(* IEC 61131-3 sources: llm-plc-st-eval/data/definitivo/gemini-3.1-pro-preview/I8/few_shot, 3 files *)

(* ---- ejec_1.st ---- *)
FUNCTION_BLOCK FB_Compresor
VAR_INPUT
    pOilOk : BOOL;    (* Presion de aceite correcta *)
    tempOk : BOOL;    (* Temperatura correcta *)
    sinAlm : BOOL;    (* Ausencia de alarmas *)
    btnMarcha : BOOL; (* Boton de arranque *)
    btnParo : BOOL;   (* Boton de parada *)
END_VAR
VAR_OUTPUT
    comp : BOOL;      (* Salida del compresor *)
    causaBloqueo : INT; (* Causa de bloqueo: 1=Aceite, 2=Temp, 3=Alarma, 0=Ninguno *)
END_VAR
VAR
    tonOil : TON;     (* Temporizador para presion de aceite *)
    trigMarcha : R_TRIG; (* Detector de flanco para boton de marcha *)
    permisivosOk : BOOL; (* Estado de todos los permisivos *)
END_VAR

(* Temporizador: presion de aceite activa por 3 segundos continuos *)
tonOil(IN := pOilOk, PT := T#3S);

(* Determinacion de la causa de bloqueo con prioridad (menor numero primero) *)
IF NOT tonOil.Q THEN
    causaBloqueo := 1;
ELSIF NOT tempOk THEN
    causaBloqueo := 2;
ELSIF NOT sinAlm THEN
    causaBloqueo := 3;
ELSE
    causaBloqueo := 0;
END_IF;

(* Evaluacion global de permisivos *)
permisivosOk := (causaBloqueo = 0);

(* Deteccion de flanco de subida del boton de marcha *)
trigMarcha(CLK := btnMarcha);

(* Logica de control del compresor (Paro prioritario y perdida de permisivos) *)
IF btnParo OR NOT permisivosOk THEN
    comp := FALSE;
ELSIF trigMarcha.Q AND permisivosOk THEN
    comp := TRUE;
END_IF;
END_FUNCTION_BLOCK

(* ---- ejec_2.st ---- *)
FUNCTION_BLOCK FB_Compresor
VAR_INPUT
    pOilOk : BOOL; (* Presion de aceite *)
    tempOk : BOOL; (* Temperatura correcta *)
    sinAlm : BOOL; (* Ausencia de alarmas *)
    btnMarcha : BOOL; (* Boton de arranque *)
    btnParo : BOOL; (* Boton de parada *)
END_VAR
VAR_OUTPUT
    comp : BOOL; (* Mando del compresor *)
    causaBloqueo : INT; (* Codigo de permisivo faltante *)
END_VAR
VAR
    tOil : TON; (* Temporizador de presion de aceite *)
    trigMarcha : R_TRIG; (* Detector de flanco de marcha *)
    permisivosOk : BOOL; (* Estado de todos los permisivos *)
END_VAR

(* Temporizador para validar la presion de aceite por 3s continuos *)
tOil(IN := pOilOk, PT := T#3S);

(* Deteccion de flanco de subida del boton de marcha *)
trigMarcha(CLK := btnMarcha);

(* Evaluacion general de permisivos *)
permisivosOk := tOil.Q AND tempOk AND sinAlm;

(* Logica de arranque y parada (prioridad al paro y a la perdida de permisivos) *)
IF btnParo OR NOT permisivosOk THEN
    comp := FALSE;
ELSIF trigMarcha.Q AND permisivosOk THEN
    comp := TRUE;
END_IF;

(* Determinacion de la causa de bloqueo (prioridad al numero menor) *)
IF NOT tOil.Q THEN
    causaBloqueo := 1; (* Falta presion de aceite *)
ELSIF NOT tempOk THEN
    causaBloqueo := 2; (* Falta temperatura correcta *)
ELSIF NOT sinAlm THEN
    causaBloqueo := 3; (* Alarma activa *)
ELSE
    causaBloqueo := 0; (* Todos los permisivos OK *)
END_IF;
END_FUNCTION_BLOCK

(* ---- ejec_3.st ---- *)
FUNCTION_BLOCK FB_Compresor
VAR_INPUT
    pOilOk : BOOL;    (* Presion de aceite correcta *)
    tempOk : BOOL;    (* Temperatura correcta *)
    sinAlm : BOOL;    (* Ausencia de alarmas *)
    btnMarcha : BOOL; (* Boton de arranque *)
    btnParo : BOOL;   (* Boton de parada *)
END_VAR
VAR_OUTPUT
    comp : BOOL;        (* Mando del compresor *)
    causaBloqueo : INT; (* Codigo de permisivo faltante *)
END_VAR
VAR
    tOil : TON;           (* Temporizador de presion de aceite *)
    trigMarcha : R_TRIG;  (* Detector de flanco para el arranque *)
    permisivosOk : BOOL;  (* Estado global de permisivos *)
END_VAR

(* Validacion de presion de aceite continua por 3 segundos *)
tOil(IN := pOilOk, PT := T#3S);

(* Determinacion de la causa de bloqueo (prioridad al numero menor) *)
IF NOT tOil.Q THEN
    causaBloqueo := 1;
ELSIF NOT tempOk THEN
    causaBloqueo := 2;
ELSIF NOT sinAlm THEN
    causaBloqueo := 3;
ELSE
    causaBloqueo := 0;
END_IF;

(* Todos los permisivos se cumplen si no hay causa de bloqueo *)
permisivosOk := (causaBloqueo = 0);

(* Deteccion de pulsacion del boton de marcha (transicion FALSE a TRUE) *)
trigMarcha(CLK := btnMarcha);

(* Control de marcha y paro del compresor (Paro prioritario) *)
IF btnParo OR NOT permisivosOk THEN
    comp := FALSE;
ELSIF trigMarcha.Q THEN
    comp := TRUE;
END_IF;
END_FUNCTION_BLOCK
